FUNCTION_BLOCK FB_OpenClose_Vlave
VAR_INPUT
	val_AfterPump	: E_Pis_Name;
	Pump_ID			: E_Pump_List:=E_Pump_List.eNotSelected;
END_VAR
VAR_OUTPUT
END_VAR
VAR
	stPist	: REFERENCE TO ST_Piston;
	stPump	: REFERENCE TO ST_Pump	;
	bOneTime	:	BOOL	;
END_VAR

act_SetReference();

IF (stPump.bRun_Auto OR stPump.bRun_Man) THEN
	bOneTime:=FALSE;
	IF NOT stPist.st_Open THEN
		stPist.req_Open:=TRUE;
	END_IF
ELSE
	IF NOT stPist.st_Close AND NOT bOneTime THEN
		stPist.req_Close:=TRUE;
		bOneTime:=TRUE;
	END_IF
END_IF

ACTION act_SetReference:
stPist REF= stPis[val_AfterPump];
stPump REF= g_Pump.arr_st_Pump[Pump_ID];
END_ACTION

END_FUNCTION_BLOCK

(* stored: Version 1.1.0.1, ProductVersion 3.1.4024.12
   POU FB_OpenClose_Vlave: Id {ee22d19d-71e8-4576-8a06-4d683eae0d16}, SpecialFunc None
   Action act_SetReference: Id {ffb6f6bd-25a2-4260-b172-60c0ca3a9d6f} *)
